Fanuc KAREL source: KO00130.KL

PROGRAM KO00130
%NOLOCKGROUP
VAR
  R: REAL
  CFG: CONFIG
  OUT: XYZWPR
  N: REAL
BEGIN
  N = 1
  R = 2.0
  CFG.CFG_FLIP = TRUE
  OUT = POS(N, R, R, R, R, R, CFG)
END KO00130
